DATA_BLOCK "FRK_PersistRootSince"
{ S7_Optimized_Access := 'TRUE' }
VERSION : 0.1
NON_RETAIN
VAR
    SinceMs {ExternalAccessible := 'False'; ExternalVisible := 'False'; ExternalWritable := 'False'} : Array[1..1] of UDInt;
    WasPending {ExternalAccessible := 'False'; ExternalVisible := 'False'; ExternalWritable := 'False'} : Array[1..1] of Bool;
END_VAR
BEGIN
END_DATA_BLOCK
